Fanuc KAREL source: KB00016.KL

PROGRAM KB00016
%NOLOCKGROUP
%ENVIRONMENT BYNAM
VAR
  P1: STRING[80]
  P2: INTEGER
  P3: INTEGER
  P4: BOOLEAN
BEGIN
  P1 = 'A'
  P2 = 1
  P3 = 1
  P4 = TRUE
  CALL_PROGLIN(P1, P2, P3, P4)
END KB00016
